PROGRAM main
  VAR
    S1 AT %IX0.0  : BOOL; (* marcha, NA *)
    S0 AT %IX0.1  : BOOL; (* parada, NC: TRUE sin pulsar *)
    KM1 AT %QX0.0 : BOOL; (* línea *)
    KM2 AT %QX0.1 : BOOL; (* estrella *)
    KM3 AT %QX0.2 : BOOL; (* triángulo *)
    H1 AT %QX0.3  : BOOL; (* piloto en marcha *)
    ETAPA         : INT; (* 0 parado, 1 estrella, 2 pausa, 3 triángulo *)
    T_EST         : TON;
    T_PAU         : TON;
    FIN_EST       : BOOL;
    FIN_PAU       : BOOL;
    E0            : BOOL; (* ETAPA = 0 *)
    E1            : BOOL; (* ETAPA = 1 *)
    E2            : BOOL; (* ETAPA = 2 *)
    E3            : BOOL; (* ETAPA = 3 *)
  END_VAR
  VAR  (* added by the conversion: wires and edge detectors of the diagram *)
    _EQ1_OUT : BOOL;
    _EQ5_OUT : BOOL;
    _EQ9_OUT : BOOL;
    _AND18_OUT : BOOL;
    _SEL17_OUT : INT;
    _AND26_OUT : BOOL;
    _SEL25_OUT : INT;
    _NOT33_OUT : BOOL;
    _SEL32_OUT : INT;
    _NOT38_OUT : BOOL;
  END_VAR

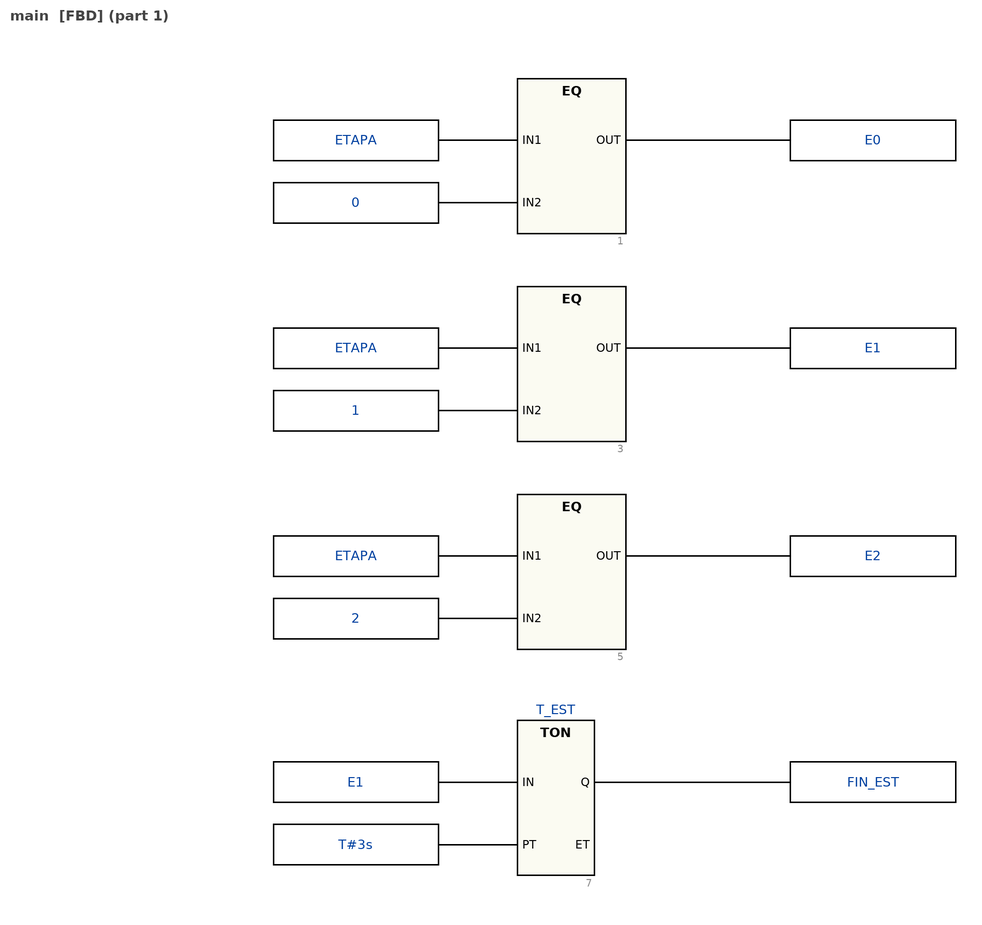
(* FBD diagram, written out as Structured Text *)
_EQ1_OUT := ETAPA = 0;
E0 := _EQ1_OUT;
_EQ5_OUT := ETAPA = 1;
E1 := _EQ5_OUT;
_EQ9_OUT := ETAPA = 2;
E2 := _EQ9_OUT;
T_EST(IN := E1, PT := T#3s);
FIN_EST := T_EST.Q;
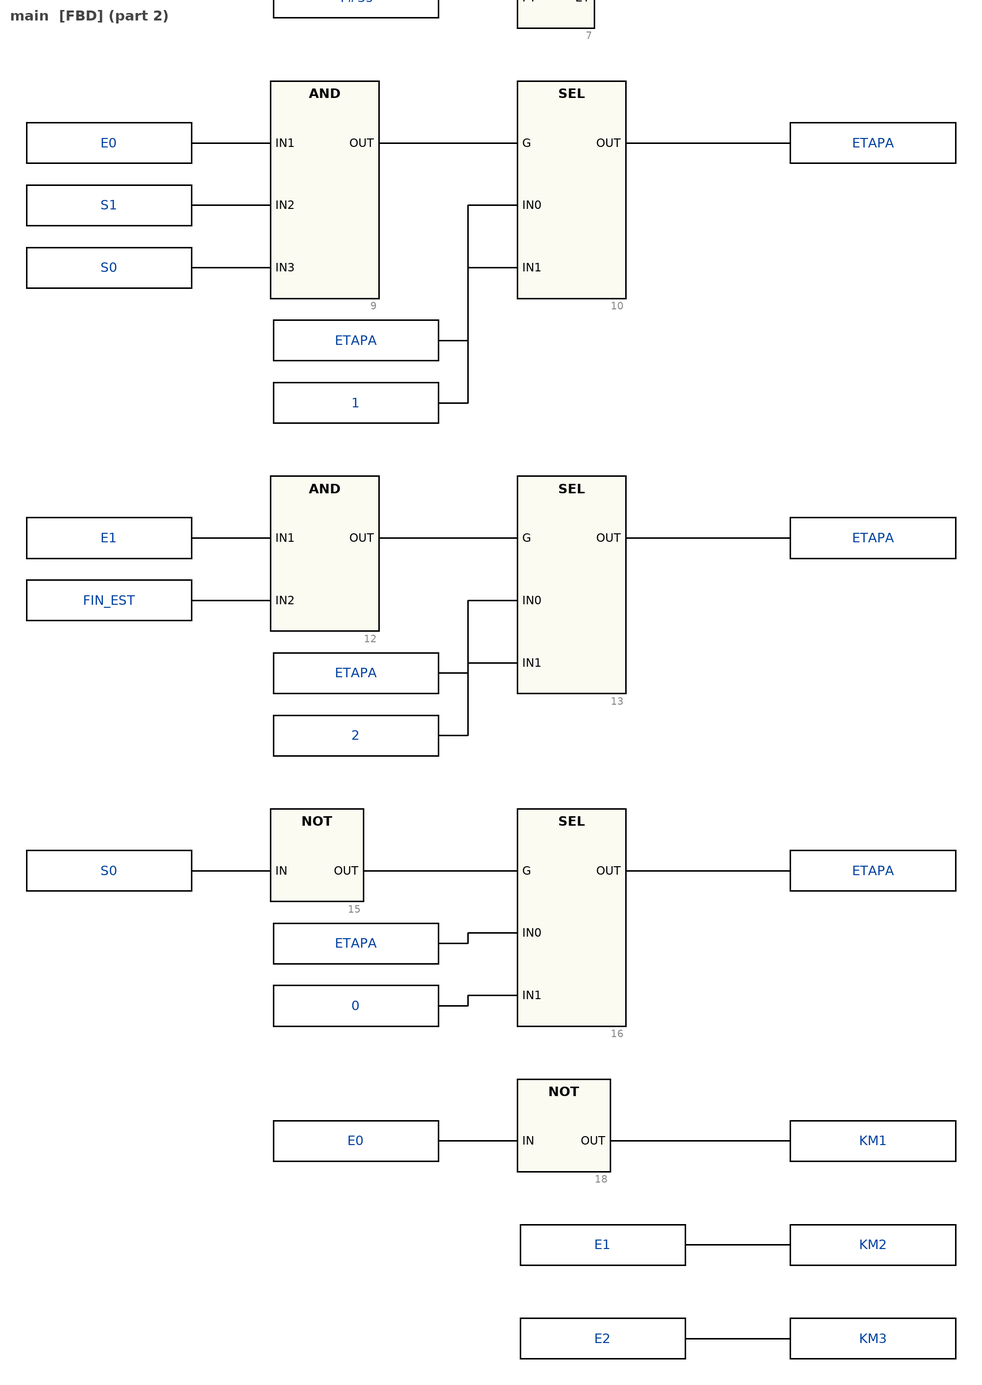
_AND18_OUT := E0 AND S1 AND S0;
_SEL17_OUT := SEL(_AND18_OUT, ETAPA, 1);
ETAPA := _SEL17_OUT;
_AND26_OUT := E1 AND FIN_EST;
_SEL25_OUT := SEL(_AND26_OUT, ETAPA, 2);
ETAPA := _SEL25_OUT;
_NOT33_OUT := NOT S0;
_SEL32_OUT := SEL(_NOT33_OUT, ETAPA, 0);
ETAPA := _SEL32_OUT;
_NOT38_OUT := NOT E0;
KM1 := _NOT38_OUT;
KM2 := E1;
KM3 := E2;
END_PROGRAM
